Omron CX-Programmer project NewProject (CX-Programmer 9.61)

# PLC NewPLC1: CJ1M CPU21

## Program Probe (cyclic task 0)

### Section Section1

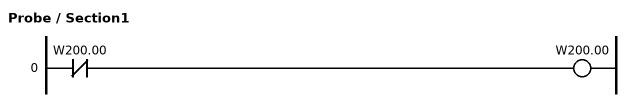
; rung 0
LDNOT W200.00
OUT W200.00

### Section END
; rung 0
END(001)